(* IEC 61131-3 sources: volt/packages/volt-lsp-iec/test-corpus/pro2193/Device/Plc Logic/Application/99 Library/Function Blocks/Alarms, 3 files *)

(* ---- enumErrorReaction.dut ---- *)
{attribute 'qualified_only'}
{attribute 'strict'}
TYPE enumErrorReaction :
(
	No_reaction		:= TO_WORD(L_IE1P.L_IE1P_Reaction.No_Reaction),	// No reaction, cycle continues
	EndCycle		:= TO_WORD(L_IE1P.L_IE1P_Reaction.CycleStop),	// Switch to 'Completing' state
	Stop			:= TO_WORD(L_IE1P.L_IE1P_Reaction.NormalStop),	// Switch to 'Stopping' state
	FastStop		:= TO_WORD(L_IE1P.L_IE1P_Reaction.FastStop)		// Switch to 'Aborting' state
) WORD;
END_TYPE

// Subset of Lenze enum: L_IE1P.L_IE1P_Reaction

// If needed we can use L_IE1P_Reaction.UserReaction1 & 2 & 6, I don't think we need this.

(* ---- enumErrorSeverity.dut ---- *)
{attribute 'qualified_only'}
{attribute 'strict'}
TYPE enumErrorSeverity :
(
	No_response		:= TO_USINT(L_IE1P.L_IE1P_SeverityLevel.No_Response),	// No reaction
	Warning			:= TO_USINT(L_IE1P.L_IE1P_SeverityLevel.Warning),		// No acknowledgement
	Information		:= TO_USINT(L_IE1P.L_IE1P_SeverityLevel.Information),	// No acknowledgement
	Warning_Lock	:= TO_USINT(L_IE1P.L_IE1P_SeverityLevel.Warning_Lock),	// Needs acknowledgement
	Fault			:= TO_USINT(L_IE1P.L_IE1P_SeverityLevel.Fault)			// Needs acknowledgement
) USINT;
END_TYPE

// Subset of Lenze enum: L_IE1P.L_IE1P_SeverityLevel

(* ---- SetErrorFB.pou ---- *)
{attribute 'monitoring_display' := 'active'}
FUNCTION_BLOCK PUBLIC SetErrorFB
VAR_INPUT
	moduleHandler	: L_IMHP.L_IMHP_IModuleHandler;
	textRefId		: WORD;				// Id of error-textlist
	errorId			: WORD;				// Id of error in the error-textlist
	alarmCondition	: BOOL;				// Condition to set the alarm.
	alarmDelay		: REAL;				// Time after which the alarm trips (in sec.)
	severity		: enumErrorSeverity := enumErrorSeverity.Fault;
	reaction		: enumErrorReaction := enumErrorReaction.No_reaction;
	testAlarm		: BOOL;
END_VAR
VAR_OUTPUT
	active			: BOOL;				// Alarm is active.
END_VAR
VAR
	SetErrorSingle	: L_IE1P.L_IE1P_SetErrorSingle;
	AlarmTimeout	: BTON;

	KeepShittyAlarmHigh : Standard.TOF;	// todo: test if this is still needed!!
END_VAR

%LANGUAGE CFC UNSUPPORTED

END_FUNCTION_BLOCK

METHOD PRIVATE CheckRefs

%LANGUAGE ST
IF moduleHandler = 0 THEN
	ThrowException('No modulehandler for SetErrorFB');
END_IF

IF textRefId = 0 THEN
	ThrowException('No textrefid for SetErrorFB');
END_IF

IF SetErrorSingle.xSetError AND textRefId <> 15372 AND textRefId <> 15373 AND textRefId <> 15374 THEN
	GlobalVars.activeAlarmInstance		:= CONCAT3(DWORD_TO_HEXSTRING(textRefId),':',TO_STRING(errorId));
END_IF

END_METHOD

METHOD PRIVATE ConvertSeverityAndReaction

%LANGUAGE ST
{warning disable C0327}	// Implicit conversion from one enumeration type to another.
SetErrorSingle.eReaction		:= reaction;
SetErrorSingle.eSeverity		:= severity;
{warning restore C0327}	// Implicit conversion from one enumeration type to another.

END_METHOD

// Get the elapsed time of the alarm timer.
{attribute 'monitoring':='call'}
PROPERTY PUBLIC ElapsedTime : REAL

GET
VAR
END_VAR

%LANGUAGE ST
IF AlarmTimeout.TON1.IN THEN
	ElapsedTime := TO_REAL(AlarmTimeout.TON1.ET) / 1000;
END_IF

END_GET
END_PROPERTY
